(* PLC project canworks, canworks canworks-deploy VERSION *)
(* stored: creationDateTime 2026-10-23T00:00:00 *)
(* canworks PLC link for canworks-bridge: Modbus TCP port 1502, unit 1, word order high_first, map hash 16#8BFA51BC. Generated by canworks-deploy VERSION; export again after a config change. *)

(* canworks values; generated, export again after a config change *)
TYPE canworks_values : STRUCT
  ok : BOOL;  (* canworks-bridge answers and serves this program's map *)
  bus_ok : BOOL;  (* ok, and every CAN network of the bridge has its bus up (status byte 7 bit 1 clear) *)
  link : ARRAY[0..1279] OF WORD;  (* the bridge's control, SDO, live list and mailbox words: the canworks blocks' LINK *)
  in_w : ARRAY[0..259] OF WORD;  (* input registers 0..259, read with function 4 *)
  out_w : ARRAY[0..94] OF WORD;  (* holding registers 0..94, written with function 16 *)
  can_bus_state : USINT;  (* CAN bus state *)
  can_master_state : USINT;  (* CANopen master state *)
  rtd_ok : BOOL;  (* node rtd (5): operational *)
  rtd_state : USINT;  (* node rtd (5): NMT state *)
  rtd_emcy : WORD;  (* node rtd (5): last EMCY code *)
  rtd_tpdo1_timeout : BOOL;  (* node rtd (5): TPDO 1 receive timeout *)
  rtd_AI0_Input_PV : INT;  (* node rtd (5) TPDO1 0x7130:1 AI0_Input_PV *)
  rtd_AI1_Input_PV : INT;  (* node rtd (5) TPDO1 0x7130:2 AI1_Input_PV *)
  rtd_AI2_Input_PV : INT;  (* node rtd (5) TPDO1 0x7130:3 AI2_Input_PV *)
  rtd_AI3_Input_PV : INT;  (* node rtd (5) TPDO1 0x7130:4 AI3_Input_PV *)
  dio_ok : BOOL;  (* node dio (6): operational *)
  dio_state : USINT;  (* node dio (6): NMT state *)
  dio_emcy : WORD;  (* node dio (6): last EMCY code *)
  dio_Read_input_8_bit_1 : USINT;  (* node dio (6) TPDO1 0x6000:1 Read input 8-bit 1 *)
  dio_Read_input_8_bit_2 : USINT;  (* node dio (6) TPDO1 0x6000:2 Read input 8-bit 2 *)
  dio_Read_analogue_input_1 : INT;  (* node dio (6) TPDO1 0x6401:1 Read analogue input 1 *)
  dio_Read_analogue_input_2 : INT;  (* node dio (6) TPDO1 0x6401:2 Read analogue input 2 *)
  dio_Write_output_8_bit_1 : USINT;  (* node dio (6) RPDO1 0x6200:1 Write output 8-bit 1 *)
  dio_Write_output_8_bit_2 : USINT;  (* node dio (6) RPDO1 0x6200:2 Write output 8-bit 2 *)
  dio_Write_analogue_output_1 : INT;  (* node dio (6) RPDO1 0x6411:1 Write analogue output 1 *)
  dio_Write_analogue_output_2 : INT;  (* node dio (6) RPDO1 0x6411:2 Write analogue output 2 *)
END_STRUCT;
END_TYPE

PROGRAM canworks_in
  VAR_EXTERNAL
    canworks : canworks_values;
  END_VAR
  VAR
    last_counter : WORD;
    moved : BOOL;
    stale : TON;
    link_service : CW_LINK_SERVICE;
  END_VAR

(* Generated by canworks: do not edit, export the map again after a config change. *)
moved := canworks.in_w[3] <> last_counter;
last_counter := canworks.in_w[3];
stale(IN := NOT moved, PT := T#3000ms);
canworks.ok := canworks.in_w[0] = WORD#16#8BFA AND canworks.in_w[1] = WORD#16#51BC AND NOT stale.Q;
canworks.bus_ok := canworks.ok AND (canworks.in_w[5] AND WORD#16#0002) = WORD#0;
canworks.link[21] := WORD#16#0106 OR SEL(canworks.ok, WORD#0, WORD#1);
canworks.link[0] := canworks.in_w[2];
canworks.link[1] := canworks.in_w[3];
canworks.link[2] := canworks.in_w[4];
canworks.link[3] := canworks.in_w[5];
canworks.link[14] := canworks.in_w[26];
canworks.link[15] := canworks.in_w[27];
canworks.link[16] := canworks.in_w[28];
canworks.link[17] := canworks.in_w[29];
canworks.link[18] := canworks.in_w[30];
canworks.link[19] := canworks.in_w[31];
canworks.link[20] := canworks.in_w[32];
canworks.link[25] := canworks.in_w[18];
canworks.link[26] := canworks.in_w[19];
canworks.link[27] := canworks.in_w[20];
canworks.link[28] := canworks.in_w[21];
canworks.link[29] := canworks.in_w[22];
canworks.link[30] := canworks.in_w[23];
canworks.link[31] := canworks.in_w[24];
canworks.link[32] := canworks.in_w[25];
canworks.link[89] := WORD#16#0431;
canworks.link[216] := canworks.in_w[33];
canworks.link[217] := canworks.in_w[34];
canworks.link[218] := canworks.in_w[35];
canworks.link[219] := canworks.in_w[36];
canworks.link[220] := canworks.in_w[37];
canworks.link[221] := canworks.in_w[38];
canworks.link[222] := canworks.in_w[39];
canworks.link[223] := canworks.in_w[40];
canworks.link[224] := canworks.in_w[41];
canworks.link[225] := canworks.in_w[42];
canworks.link[226] := canworks.in_w[43];
canworks.link[227] := canworks.in_w[44];
canworks.link[228] := canworks.in_w[45];
canworks.link[229] := canworks.in_w[46];
canworks.link[230] := canworks.in_w[47];
canworks.link[231] := canworks.in_w[48];
canworks.link[232] := canworks.in_w[49];
canworks.link[233] := canworks.in_w[50];
canworks.link[234] := canworks.in_w[51];
canworks.link[235] := canworks.in_w[52];
canworks.link[236] := canworks.in_w[53];
canworks.link[237] := canworks.in_w[54];
canworks.link[238] := canworks.in_w[55];
canworks.link[239] := canworks.in_w[56];
canworks.link[240] := canworks.in_w[57];
canworks.link[241] := canworks.in_w[58];
canworks.link[242] := canworks.in_w[59];
canworks.link[243] := canworks.in_w[60];
canworks.link[244] := canworks.in_w[61];
canworks.link[245] := canworks.in_w[62];
canworks.link[246] := canworks.in_w[63];
canworks.link[247] := canworks.in_w[64];
canworks.link[248] := canworks.in_w[65];
canworks.link[249] := canworks.in_w[66];
canworks.link[250] := canworks.in_w[67];
canworks.link[251] := canworks.in_w[68];
canworks.link[252] := canworks.in_w[69];
canworks.link[253] := canworks.in_w[70];
canworks.link[254] := canworks.in_w[71];
canworks.link[255] := canworks.in_w[72];
canworks.link[256] := canworks.in_w[73];
canworks.link[257] := canworks.in_w[74];
canworks.link[258] := canworks.in_w[75];
canworks.link[259] := canworks.in_w[76];
canworks.link[260] := canworks.in_w[77];
canworks.link[261] := canworks.in_w[78];
canworks.link[262] := canworks.in_w[79];
canworks.link[263] := canworks.in_w[80];
canworks.link[264] := canworks.in_w[81];
canworks.link[265] := canworks.in_w[82];
canworks.link[266] := canworks.in_w[83];
canworks.link[267] := canworks.in_w[84];
canworks.link[268] := canworks.in_w[85];
canworks.link[269] := canworks.in_w[86];
canworks.link[270] := canworks.in_w[87];
canworks.link[271] := canworks.in_w[88];
canworks.link[272] := canworks.in_w[89];
canworks.link[273] := canworks.in_w[90];
canworks.link[274] := canworks.in_w[91];
canworks.link[275] := canworks.in_w[92];
canworks.link[276] := canworks.in_w[93];
canworks.link[277] := canworks.in_w[94];
canworks.link[278] := canworks.in_w[95];
canworks.link[279] := canworks.in_w[96];
canworks.link[280] := canworks.in_w[97];
canworks.link[281] := canworks.in_w[98];
canworks.link[282] := canworks.in_w[99];
canworks.link[283] := canworks.in_w[100];
canworks.link[284] := canworks.in_w[101];
canworks.link[285] := canworks.in_w[102];
canworks.link[286] := canworks.in_w[103];
canworks.link[287] := canworks.in_w[104];
canworks.link[720] := canworks.in_w[105];
canworks.link[721] := canworks.in_w[106];
canworks.link[722] := canworks.in_w[107];
canworks.link[723] := canworks.in_w[108];
canworks.link[724] := canworks.in_w[109];
canworks.link[725] := canworks.in_w[110];
canworks.link[726] := canworks.in_w[111];
canworks.link[727] := canworks.in_w[112];
canworks.link[728] := canworks.in_w[113];
canworks.link[729] := canworks.in_w[114];
canworks.link[730] := canworks.in_w[115];
canworks.link[731] := canworks.in_w[116];
canworks.link[732] := canworks.in_w[117];
canworks.link[733] := canworks.in_w[118];
canworks.link[734] := canworks.in_w[119];
canworks.link[735] := canworks.in_w[120];
canworks.link[736] := canworks.in_w[121];
canworks.link[737] := canworks.in_w[122];
canworks.link[738] := canworks.in_w[123];
canworks.link[739] := canworks.in_w[124];
canworks.link[740] := canworks.in_w[125];
canworks.link[741] := canworks.in_w[126];
canworks.link[742] := canworks.in_w[127];
canworks.link[743] := canworks.in_w[128];
canworks.link[744] := canworks.in_w[129];
canworks.link[745] := canworks.in_w[130];
canworks.link[746] := canworks.in_w[131];
canworks.link[747] := canworks.in_w[132];
canworks.link[748] := canworks.in_w[133];
canworks.link[749] := canworks.in_w[134];
canworks.link[750] := canworks.in_w[135];
canworks.link[751] := canworks.in_w[136];
canworks.link[752] := canworks.in_w[137];
canworks.link[753] := canworks.in_w[138];
canworks.link[754] := canworks.in_w[139];
canworks.link[755] := canworks.in_w[140];
canworks.link[756] := canworks.in_w[141];
canworks.link[757] := canworks.in_w[142];
canworks.link[758] := canworks.in_w[143];
canworks.link[759] := canworks.in_w[144];
canworks.link[760] := canworks.in_w[145];
canworks.link[761] := canworks.in_w[146];
canworks.link[762] := canworks.in_w[147];
canworks.link[763] := canworks.in_w[148];
canworks.link[764] := canworks.in_w[149];
canworks.link[765] := canworks.in_w[150];
canworks.link[766] := canworks.in_w[151];
canworks.link[767] := canworks.in_w[152];
canworks.link[768] := canworks.in_w[153];
canworks.link[769] := canworks.in_w[154];
canworks.link[770] := canworks.in_w[155];
canworks.link[771] := canworks.in_w[156];
canworks.link[772] := canworks.in_w[157];
canworks.link[773] := canworks.in_w[158];
canworks.link[774] := canworks.in_w[159];
canworks.link[775] := canworks.in_w[160];
canworks.link[776] := canworks.in_w[161];
canworks.link[777] := canworks.in_w[162];
canworks.link[778] := canworks.in_w[163];
canworks.link[779] := canworks.in_w[164];
canworks.link[780] := canworks.in_w[165];
canworks.link[781] := canworks.in_w[166];
canworks.link[782] := canworks.in_w[167];
canworks.link[783] := canworks.in_w[168];
canworks.link[784] := canworks.in_w[169];
canworks.link[785] := canworks.in_w[170];
canworks.link[786] := canworks.in_w[171];
canworks.link[787] := canworks.in_w[172];
canworks.link[788] := canworks.in_w[173];
canworks.link[789] := canworks.in_w[174];
canworks.link[790] := canworks.in_w[175];
canworks.link[791] := canworks.in_w[176];
canworks.link[792] := canworks.in_w[177];
canworks.link[793] := canworks.in_w[178];
canworks.link[794] := canworks.in_w[179];
canworks.link[795] := canworks.in_w[180];
canworks.link[796] := canworks.in_w[181];
canworks.link[797] := canworks.in_w[182];
canworks.link[798] := canworks.in_w[183];
canworks.link[799] := canworks.in_w[184];
canworks.link[800] := canworks.in_w[185];
canworks.link[801] := canworks.in_w[186];
canworks.link[802] := canworks.in_w[187];
canworks.link[803] := canworks.in_w[188];
canworks.link[804] := canworks.in_w[189];
canworks.link[805] := canworks.in_w[190];
canworks.link[806] := canworks.in_w[191];
canworks.link[807] := canworks.in_w[192];
canworks.link[808] := canworks.in_w[193];
canworks.link[809] := canworks.in_w[194];
canworks.link[810] := canworks.in_w[195];
canworks.link[811] := canworks.in_w[196];
canworks.link[812] := canworks.in_w[197];
canworks.link[813] := canworks.in_w[198];
canworks.link[814] := canworks.in_w[199];
canworks.link[815] := canworks.in_w[200];
canworks.link[816] := canworks.in_w[201];
canworks.link[817] := canworks.in_w[202];
canworks.link[818] := canworks.in_w[203];
canworks.link[819] := canworks.in_w[204];
canworks.link[820] := canworks.in_w[205];
canworks.link[821] := canworks.in_w[206];
canworks.link[822] := canworks.in_w[207];
canworks.link[823] := canworks.in_w[208];
canworks.link[824] := canworks.in_w[209];
canworks.link[825] := canworks.in_w[210];
canworks.link[826] := canworks.in_w[211];
canworks.link[827] := canworks.in_w[212];
canworks.link[828] := canworks.in_w[213];
canworks.link[829] := canworks.in_w[214];
canworks.link[830] := canworks.in_w[215];
canworks.link[831] := canworks.in_w[216];
canworks.link[832] := canworks.in_w[217];
canworks.link[833] := canworks.in_w[218];
canworks.link[834] := canworks.in_w[219];
canworks.link[835] := canworks.in_w[220];
canworks.link[836] := canworks.in_w[221];
canworks.link[837] := canworks.in_w[222];
canworks.link[838] := canworks.in_w[223];
canworks.link[839] := canworks.in_w[224];
canworks.link[960] := canworks.in_w[225];
canworks.link[961] := canworks.in_w[226];
canworks.link[962] := canworks.in_w[227];
canworks.link[963] := canworks.in_w[228];
canworks.link[964] := canworks.in_w[229];
canworks.link[965] := canworks.in_w[230];
canworks.link[966] := canworks.in_w[231];
canworks.link[967] := canworks.in_w[232];
canworks.link[968] := canworks.in_w[233];
canworks.link[969] := canworks.in_w[234];
canworks.link[970] := canworks.in_w[235];
canworks.link[971] := canworks.in_w[236];
canworks.link[972] := canworks.in_w[237];
canworks.link[973] := canworks.in_w[238];
canworks.link[974] := canworks.in_w[239];
canworks.link[975] := canworks.in_w[240];
canworks.link[976] := canworks.in_w[241];
canworks.link[977] := canworks.in_w[242];
canworks.link[1104] := canworks.in_w[243];
canworks.link[1105] := canworks.in_w[244];
canworks.link[1106] := canworks.in_w[245];
canworks.link[1107] := canworks.in_w[246];
canworks.link[1108] := canworks.in_w[247];
canworks.link[1109] := canworks.in_w[248];
canworks.link[1110] := canworks.in_w[249];
canworks.link[1111] := canworks.in_w[250];
canworks.link[1112] := canworks.in_w[251];
canworks.link[1113] := canworks.in_w[252];
canworks.link[1114] := canworks.in_w[253];
canworks.link[1115] := canworks.in_w[254];
canworks.link[1116] := canworks.in_w[255];
canworks.link[1117] := canworks.in_w[256];
canworks.link[1118] := canworks.in_w[257];
canworks.link[1119] := canworks.in_w[258];
canworks.link[1120] := canworks.in_w[259];
link_service(LINK := canworks.link);
canworks.can_bus_state := SEL(canworks.ok, USINT#0, WORD_TO_USINT((canworks.in_w[13] AND WORD#16#00FF)));
canworks.can_master_state := SEL(canworks.ok, USINT#0, WORD_TO_USINT(SHR(canworks.in_w[13], 8)));
canworks.rtd_ok := SEL(canworks.ok, FALSE, (canworks.in_w[14] AND WORD#16#0100) <> WORD#0);
canworks.rtd_state := SEL(canworks.ok, USINT#0, WORD_TO_USINT((canworks.in_w[14] AND WORD#16#00FF)));
canworks.rtd_emcy := SEL(canworks.ok, WORD#0, canworks.in_w[16]);
canworks.rtd_tpdo1_timeout := SEL(canworks.ok, FALSE, (canworks.in_w[14] AND WORD#16#0400) <> WORD#0);
canworks.rtd_AI0_Input_PV := WORD_TO_INT(canworks.in_w[6]);
canworks.rtd_AI1_Input_PV := WORD_TO_INT(canworks.in_w[7]);
canworks.rtd_AI2_Input_PV := WORD_TO_INT(canworks.in_w[8]);
canworks.rtd_AI3_Input_PV := WORD_TO_INT(canworks.in_w[9]);
canworks.dio_ok := SEL(canworks.ok, FALSE, (canworks.in_w[14] AND WORD#16#0200) <> WORD#0);
canworks.dio_state := SEL(canworks.ok, USINT#0, WORD_TO_USINT(SHR(canworks.in_w[15], 8)));
canworks.dio_emcy := SEL(canworks.ok, WORD#0, canworks.in_w[17]);
canworks.dio_Read_input_8_bit_1 := WORD_TO_USINT(SHR(canworks.in_w[10], 8));
canworks.dio_Read_input_8_bit_2 := WORD_TO_USINT((canworks.in_w[10] AND WORD#16#00FF));
canworks.dio_Read_analogue_input_1 := WORD_TO_INT(canworks.in_w[11]);
canworks.dio_Read_analogue_input_2 := WORD_TO_INT(canworks.in_w[12]);
END_PROGRAM

PROGRAM canworks_out
  VAR_EXTERNAL
    canworks : canworks_values;
  END_VAR

(* Generated by canworks: do not edit, export the map again after a config change. *)
canworks.out_w[3] := SHL((USINT_TO_WORD(canworks.dio_Write_output_8_bit_1) AND WORD#16#00FF), 8) OR (USINT_TO_WORD(canworks.dio_Write_output_8_bit_2) AND WORD#16#00FF);
canworks.out_w[4] := INT_TO_WORD(canworks.dio_Write_analogue_output_1);
canworks.out_w[5] := INT_TO_WORD(canworks.dio_Write_analogue_output_2);
canworks.out_w[6] := canworks.link[4];
canworks.out_w[7] := canworks.link[5];
canworks.out_w[8] := canworks.link[6];
canworks.out_w[9] := canworks.link[7];
canworks.out_w[10] := canworks.link[8];
canworks.out_w[11] := canworks.link[9];
canworks.out_w[12] := canworks.link[10];
canworks.out_w[13] := canworks.link[11];
canworks.out_w[14] := canworks.link[12];
canworks.out_w[15] := canworks.link[13];
canworks.out_w[16] := canworks.link[144];
canworks.out_w[17] := canworks.link[145];
canworks.out_w[18] := canworks.link[146];
canworks.out_w[19] := canworks.link[147];
canworks.out_w[20] := canworks.link[148];
canworks.out_w[21] := canworks.link[149];
canworks.out_w[22] := canworks.link[150];
canworks.out_w[23] := canworks.link[151];
canworks.out_w[24] := canworks.link[152];
canworks.out_w[25] := canworks.link[153];
canworks.out_w[26] := canworks.link[154];
canworks.out_w[27] := canworks.link[155];
canworks.out_w[28] := canworks.link[156];
canworks.out_w[29] := canworks.link[157];
canworks.out_w[30] := canworks.link[158];
canworks.out_w[31] := canworks.link[159];
canworks.out_w[32] := canworks.link[160];
canworks.out_w[33] := canworks.link[161];
canworks.out_w[34] := canworks.link[162];
canworks.out_w[35] := canworks.link[163];
canworks.out_w[36] := canworks.link[164];
canworks.out_w[37] := canworks.link[165];
canworks.out_w[38] := canworks.link[166];
canworks.out_w[39] := canworks.link[167];
canworks.out_w[40] := canworks.link[168];
canworks.out_w[41] := canworks.link[169];
canworks.out_w[42] := canworks.link[170];
canworks.out_w[43] := canworks.link[171];
canworks.out_w[44] := canworks.link[172];
canworks.out_w[45] := canworks.link[173];
canworks.out_w[46] := canworks.link[174];
canworks.out_w[47] := canworks.link[175];
canworks.out_w[48] := canworks.link[176];
canworks.out_w[49] := canworks.link[177];
canworks.out_w[50] := canworks.link[178];
canworks.out_w[51] := canworks.link[179];
canworks.out_w[52] := canworks.link[180];
canworks.out_w[53] := canworks.link[181];
canworks.out_w[54] := canworks.link[182];
canworks.out_w[55] := canworks.link[183];
canworks.out_w[56] := canworks.link[184];
canworks.out_w[57] := canworks.link[185];
canworks.out_w[58] := canworks.link[186];
canworks.out_w[59] := canworks.link[187];
canworks.out_w[60] := canworks.link[188];
canworks.out_w[61] := canworks.link[189];
canworks.out_w[62] := canworks.link[190];
canworks.out_w[63] := canworks.link[191];
canworks.out_w[64] := canworks.link[192];
canworks.out_w[65] := canworks.link[193];
canworks.out_w[66] := canworks.link[194];
canworks.out_w[67] := canworks.link[195];
canworks.out_w[68] := canworks.link[196];
canworks.out_w[69] := canworks.link[197];
canworks.out_w[70] := canworks.link[198];
canworks.out_w[71] := canworks.link[199];
canworks.out_w[72] := canworks.link[200];
canworks.out_w[73] := canworks.link[201];
canworks.out_w[74] := canworks.link[202];
canworks.out_w[75] := canworks.link[203];
canworks.out_w[76] := canworks.link[204];
canworks.out_w[77] := canworks.link[205];
canworks.out_w[78] := canworks.link[206];
canworks.out_w[79] := canworks.link[207];
canworks.out_w[80] := canworks.link[208];
canworks.out_w[81] := canworks.link[209];
canworks.out_w[82] := canworks.link[210];
canworks.out_w[83] := canworks.link[211];
canworks.out_w[84] := canworks.link[212];
canworks.out_w[85] := canworks.link[213];
canworks.out_w[86] := canworks.link[214];
canworks.out_w[87] := canworks.link[215];
canworks.out_w[88] := canworks.link[102];
canworks.out_w[89] := canworks.link[103];
canworks.out_w[90] := canworks.link[104];
canworks.out_w[91] := canworks.link[128];
canworks.out_w[92] := canworks.link[129];
canworks.out_w[93] := canworks.link[130];
canworks.out_w[94] := canworks.link[131];
(* PLC link header, last: running, then the map hash 0x8bfa51bc *)
canworks.out_w[1] := WORD#16#8BFA;
canworks.out_w[2] := WORD#16#51BC;
canworks.out_w[0] := WORD#1;
END_PROGRAM

CONFIGURATION canworks_config
  RESOURCE canworks_res ON PLC
    VAR_GLOBAL
      canworks : canworks_values;  (* canworks values; generated, export again after a config change *)
    END_VAR
    TASK canworks_task(INTERVAL := T#200ms, PRIORITY := 1);
    PROGRAM canworks_in_instance WITH canworks_task : canworks_in;
    PROGRAM canworks_out_instance WITH canworks_task : canworks_out;
  END_RESOURCE
END_CONFIGURATION
